// TIA Portal project "stage ocp" (V17)

(* hardware
DEVICE "S7-300/ET200M station_1"  S7-300 station
   slot 0: "Rail_0"  Rail  6ES7 390-1***0-0AA0
   slot 2: "PLC_1"  CPU 315-2 DP  6ES7 315-2AH14-0AB0  V3.0
      slot 0: "MPI interface_1"  MPI
      slot 1: "DP interface_1"  DP
   slot 4: "CP 341 RS422/485_1"  CP 341 RS422/485  6ES7 341-1CH02-0AE0  V2.0
   slot 5: "CP 343-1 Lean_1"  CP 343-1 LEAN  6GK7 343-1CX10-0XE0  V3.0
   slot 6: "DI 16x24VDC_1"  DI16 x 24VDC, interrupt  6ES7 321-7BH01-0AB0
   slot 7: "DO 16x24VDC/0.5A_1"  DO16xDC24V/0.5A  6ES7 322-8BH10-0AB0
DEVICE "SCALANCE XC-100 unmanaged"  SCALANCE X-Station
   slot 0: "SCALANCE X rack"  Rail
   slot 0: "Switch_1"  6GK5 106-2BB00-2AC2  V1.0
DEVICE "HMI_2"  KTP700 Basic PN
   slot 0: "HMI_2"  KTP700 Basic PN  6AV2 123-2GB03-0AX0  17.0.0.0
   slot 1: "HMI_RT_2"  KTP700 Basic PN  6AV2 123-2GB03-0AX0  17.0.0.0
   slot 5: "HMI_2.IE_CP_1"  PROFINET Interface  17.0.0.0
      slot 1: "PROFINET Interface_1"  PROFINET Interface
         slot 1: "Port_1"  Port
*)

// ===== PLC "PLC_1"  CPU 315-2 DP =====

VAR_GLOBAL   // PLC tag table "Default tag table"
   "analog input" AT %I0.0 : Bool;
   "analog outputs" AT %Q0.5 : Bool;
END_VAR

VAR_GLOBAL   // PLC tag table "Actionneur/bouton"
   "AR" AT %M0.2 : Bool;
   "MA" AT %M0.3 : Bool;
   "K1" AT %Q0.0 : Bool;
   "M" AT %Q0.1 : Bool;
   "AT" AT %Q0.2 : Bool;
   "defaut" AT %Q0.3 : Bool;
   "detect_defaut" AT %M0.4 : Bool;
   "INSTANT" AT %M0.5 : Bool;
   "10s" AT %M0.6 : Bool;
   "15s" AT %M0.7 : Bool;
   "marche" AT %M1.0 : Bool;
END_VAR

DATA_BLOCK "DB_TeSysT_Data"   // DB1
{ S7_Optimized_Access := 'FALSE' }
VERSION : 0.1
   VAR
      MotorCurrent : Int;
      SystemStatus : Word;
      tripstatus : Word;
      faultcode : Int;
      thermalstate : Int;
      MotorRunCmd : Word;
   END_VAR
BEGIN
END_DATA_BLOCK

DATA_BLOCK "hmi communication"   // DB2
{ S7_Optimized_Access := 'FALSE' }
VERSION : 0.1
   VAR
      AR : Bool;
      MA : Bool;
      K1 : Bool;
      "M" : Bool;
      AT : Bool;
      defaut : Bool;
      detect_defaut : Bool;
   END_VAR
BEGIN
END_DATA_BLOCK

ORGANIZATION_BLOCK "Main"   // OB1, LAD
TITLE = "Main Program Sweep (Cycle)"
{ S7_Optimized_Access := 'FALSE' }
VERSION : 0.1
   VAR_TEMP
      OB1_EV_CLASS : Byte;   // Bits 0-3 = 1 (Coming event), Bits 4-7 = 1 (Event class 1)
      OB1_SCAN_1 : Byte;   // 1 (Cold restart scan 1 of OB 1), 3 (Scan 2-n of OB 1)
      OB1_PRIORITY : Byte;   // Priority of OB Execution
      OB1_OB_NUMBR : Byte;   // 1 (Organization block 1, OB1)
      OB1_RESERVED_1 : Byte;   // Reserved for system
      OB1_RESERVED_2 : Byte;   // Reserved for system
      OB1_PREV_CYCLE : Int;   // Cycle time of previous OB1 scan (milliseconds)
      OB1_MIN_CYCLE : Int;   // Minimum cycle time of OB1 (milliseconds)
      OB1_MAX_CYCLE : Int;   // Maximum cycle time of OB1 (milliseconds)
      OB1_DATE_TIME : Date_And_Time;   // Date and time OB1 started
   END_VAR
BEGIN

REGION Network 1
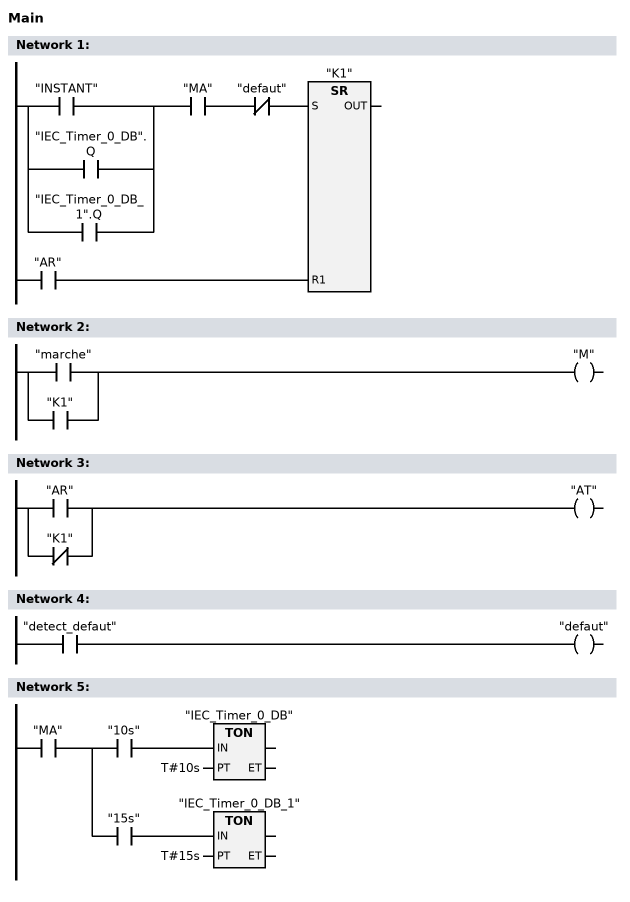
   RUNG wire#powerrail
      Contact( "INSTANT" )
      wire#w1
      Contact( "MA" )
      I_Contact( "defaut" )
      S_SR(operand := "K1", r1 := wire#w2)
   END_RUNG
   RUNG wire#powerrail
      Contact( "IEC_Timer_0_DB".Q )
   END_RUNG wire#w1
   RUNG wire#powerrail
      Contact( "IEC_Timer_0_DB_1".Q )
   END_RUNG wire#w1
   RUNG wire#powerrail
      Contact( "AR" )
   END_RUNG wire#w2
   // the same network as SCL:
   IF ("INSTANT" OR "IEC_Timer_0_DB".Q OR "IEC_Timer_0_DB_1".Q) AND "MA" AND NOT "defaut" THEN
       "K1" := TRUE;   // SR flip-flop
   END_IF;
   IF "AR" THEN "K1" := FALSE; END_IF;
END_REGION

REGION Network 2
   RUNG wire#powerrail
      Contact( "marche" )
      wire#w1
      Coil( "M" )
   END_RUNG
   RUNG wire#powerrail
      Contact( "K1" )
   END_RUNG wire#w1
   // the same network as SCL:
   "M" := "marche" OR "K1";
END_REGION

REGION Network 3
   RUNG wire#powerrail
      Contact( "AR" )
      wire#w1
      Coil( "AT" )
   END_RUNG
   RUNG wire#powerrail
      I_Contact( "K1" )
   END_RUNG wire#w1
   // the same network as SCL:
   "AT" := "AR" OR NOT "K1";
END_REGION

REGION Network 4
   RUNG wire#powerrail
      Contact( "detect_defaut" )
      Coil( "defaut" )
   END_RUNG
   // the same network as SCL:
   "defaut" := "detect_defaut";
END_REGION

REGION Network 5
   "IEC_Timer_0_DB".TON(IN := "MA" AND "10s", PT := T#10s);
   "IEC_Timer_0_DB_1".TON(IN := "MA" AND "15s", PT := T#15s);
END_REGION
END_ORGANIZATION_BLOCK

(* ===== HMI "HMI_RT_2" =====
system functions are stored by id; their names below are inferred from use
connection "HMI_Connection_1": ETHERNET, SIMATIC S7 300/400 MPI

HMI tags "Default tag table"
   "Tag_ScreenNumber" : UInt, internal
   "MA" : Bool = PLC MA AT %M0.3, 1 s
   "AR" : Bool = PLC AR AT %M0.2, 1 s
   "detect_defaut" : Bool = PLC detect_defaut AT %M0.4, 1 s
   "K1" : Bool = PLC K1 AT %Q0.0, 1 s
   "defaut" : Bool = PLC defaut AT %Q0.3, 1 s
   "10s" : Bool = PLC 10s AT %M0.6, 1 s
   "15s" : Bool = PLC 15s AT %M0.7, 1 s
   "INSTANT" : Bool = PLC INSTANT AT %M0.5, 1 s
   "marche" : Bool = PLC marche AT %M1.0, 1 s

graphic list "Graphic_list_7": 0..1 'OCP_Group.svg (2)'

graphic list "Graphic_list_4": 1 'Graphic_5'; 0 'Graphic_8'

graphic list "Graphic_list_6": 0 'Graphic_9'; 1 'Graphic_6'

graphic list "Graphic_list_1": 0..1 'transparent'

graphic list "Graphic_list_3": 0 'Graphic_1'; 1 'Graphic_2'; 2 'Graphic_3'

graphic list "Graphic_list_2": 0 'IESAAutomation_Shelter-OCP_Howden_MAROC_Im2_1'

graphic list "Graphic_list_5": 1 'Graphic_4'; 0 'Graphic_7'

recipe "MOTOR_MODE": 10S <- "10s", 15S <- "15s", INSTANT <- "INSTANT"

Template "Template_1" 800x480
   Button "Exit" at 714,429 size 71x50; TextOff 'Exit'; PictureOff "ExitRuntime_KTP700_Basic_PN_TR"; PictureOn "ExitRuntime_KTP700_Basic_PN_TR"
      on Release: StopRuntime(0)
   Button "Template_Button" at 614,429 size 71x50; TextOff 'Text'
   Button "Template_Button_1" at 514,429 size 71x50; TextOff 'Text'
   Button "Template_Button_2" at 414,429 size 71x50; TextOff 'Text'
   Button "Template_Button_3" at 314,429 size 71x50; TextOff 'Text'
   Button "Template_Button_4" at 214,429 size 71x50; TextOff 'Text'
   Button "Alarms" at 114,429 size 71x50; TextOff 'Alarms'; PictureOff "AlarmDisplay_KTP700_Basic_PN_TR"; PictureOn "AlarmDisplay_KTP700_Basic_PN_TR"
      on Release: function_ef3f5d25("Alarm window_Unacknowledged", -1)
   Button "Start screen" at 14,429 size 71x50; TextOff 'Start screen'; PictureOff "NavigateHome_KTP700_Basic_PN_TR"; PictureOn "NavigateHome_KTP700_Basic_PN_TR"
      on Release: ActivateScreen("Root screen", 0)
   SymbolicIOField "Symbolic_IO_Field_Screen" at 93,9 size 600x33; TextOff '0'; TextOn '1'; TextList "TextList_ScreenNames"
      ProcessValue <- "Tag_ScreenNumber"
      on Change: ActivateScreenByNumber("Tag_ScreenNumber", 0)
   DateTimeField "HmiScreenItemData" at 695,25 size 105x25
   DateTimeField "HmiScreenItemData_1" at 695,0 size 105x25
   GraphicView "Logo" at 0,0 size 91x51; Picture "Logo of HMI_2"

screen "Root screen" 800x480, template "Template_1"
   on GenerateScreen: SetTag("Tag_ScreenNumber", 1)
   TextField "HmiScreenItemData_1" at 80,225 size 640x25; Text 'Welcome to HMI_2 (KTP700 Basic+ PN)!'
   Button "HmiScreenItemData" at 36,87 size 159x47; TextOff 'Screen0'; PictureOff "Navigates to Screen0 for KTP700 Basic+ PN 17.0.0.0"; PictureOn "Navigates to Screen0 for KTP700 Basic+ PN 17.0.0.0"
      on Release: ActivateScreen("Screen0", 0)

screen "Screen0" 800x480, template "Template_1"
   on GenerateScreen: SetTag("Tag_ScreenNumber", 2)
   TextField "HmiScreenItemData" at 80,225 size 640x25; Text 'Screen0'
   Button "Back" at 1,52 size 159x47; TextOff 'Back'
      on Release: ActivateScreen("Root screen", 0)

screen "Screen_1" 800x480
   GraphicIOField "Graphic I/O field_2" at 0,0 size 800x480; PictureList "Graphic_list_2"
   GraphicIOField "Graphic I/O field_1" at 236,80 size 173x389; PictureList "Graphic_list_1"
   Button "Button_1" at 270,138 size 101x64; TextOff 'START'
      on Press: function_b14e0dd5("MA", 0)
   Button "Button_2" at 270,237 size 101x64; TextOff 'STOP'
      on Press: function_b14e0dd5("AR", 0)
   Button "Button_3" at 268,336 size 101x64; TextOff 'default'
      on Press: function_b14e0dd5("detect_defaut", 0)
   GraphicIOField "Graphic I/O field_3" at 21,80 size 197x389; PictureList "Graphic_list_1"
   GraphicIOField "Graphic I/O field_4" at 599,284 size 190x182; PictureList "Graphic_list_1"
   Button "Button_4" at 61,130 size 125x64; TextOff 'MODE 1'
      on Press: function_eba64363(1, U 1, 1, N)
   Button "Button_5" at 61,229 size 125x64; TextOff 'MODE 2'
      on Press: function_eba64363(1, U 2, 1, N)
   Button "Button_6" at 59,328 size 125x64; TextOff 'MODE 3'
      on Press: function_eba64363(1, U 3, 1, N)
   GraphicIOField "Graphic I/O field_5" at 618,348 size 152x100; PictureList "Graphic_list_3"; PictureOff "Graphic_1"; PictureOn "Graphic_2"
      ProcessValue <- "marche"
   TextField "Text field_1" at 618,299 size 172x29; Text 'MOTOR STATUS'
   GraphicIOField "Graphic I/O field_6" at 419,82 size 173x389; PictureList "Graphic_list_1"
   GraphicIOField "Graphic I/O field_7" at 520,385 size 59x50; PictureList "Graphic_list_6"
      ProcessValue <- "defaut"
   GraphicIOField "Graphic I/O field_8" at 520,129 size 59x56; PictureList "Graphic_list_5"; PictureOn "Graphic_4"; PictureOff "Graphic_7"
      ProcessValue <- "MA"
   GraphicIOField "Graphic I/O field_9" at 520,255 size 59x55; PictureList "Graphic_list_4"
      ProcessValue <- "AR"
   TextField "Text field_2" at 434,144 size 84x23; Text 'RUNNING'
   TextField "Text field_3" at 434,272 size 84x23; Text 'RUNNING'
   TextField "Text field_4" at 434,400 size 84x23; Text 'RUNNING'
   GraphicIOField "Graphic I/O field_10" at 693,97 size 96x71; PictureList "Graphic_list_7"
   TextField "Text field_5" at 11,29 size 184x23; Text 'service d'acceuil : MFJ'
   TextField "Text field_6" at 300,22 size 134x23; Text 'SCREEN : HOME'
   DateTimeField "Date/time field_1" at 563,20 size 219x32
*)